(* IEC 61131-3 sources: codesys-to-s7/tests/corpus/C2S7-IL/neg, 1 file *)

(* ---- input.st ---- *)
FUNCTION_BLOCK FB_I
VAR_INPUT
    a : BOOL;
    b : BOOL;
END_VAR
VAR_OUTPUT
    q : BOOL;
END_VAR
q := a AND b;
END_FUNCTION_BLOCK
